(*
SPDX-FileCopyrightText: © 2026 Oleksandr Tiutyk <trofimich@gmail.com>
SPDX-License-Identifier: MIT
License: https://opensource.org/license/mit
*)

(*!
<summary>
Defines a loop composite activity that repeats its body activity while its Condition evaluates to TRUE.
</summary>
*)

INTERFACE IWhileActivity EXTENDS IExclusiveCompositeActivity

(*!
<summary>Returns the body activity executed by this loop, or 0 when no body is configured.</summary>
*)
{attribute 'monitoring' := 'call'}
PROPERTY Body : IActivity
GET
END_GET
END_PROPERTY

(*!
<summary>Returns the loop continuation condition configured for this activity.</summary>
*)
{attribute 'monitoring' := 'call'}
PROPERTY Condition : ICondition
GET
END_GET
END_PROPERTY

(*!
<summary>Configures the required loop condition and optional body activity.</summary>
<description>
Permitted only in PASSIVE_READY. Condition is required; body is optional (when 0, evaluates condition
cyclically without advancing a body activity). Assigns THIS^ as ParentActivity of supplied elements.
</description>
<param name="condition">Condition evaluated before each iteration.</param>
<param name="body">Activity executed repeatedly while condition evaluates to TRUE, or 0.</param>
*)
METHOD Configure
VAR_INPUT
	condition : ICondition;
	body : IActivity;
END_VAR
END_METHOD

END_INTERFACE

(* stored: Version 1.1.0.1
   Itf IWhileActivity: Id {48afd1de-38c9-486e-a527-23b68379f379}
   Property Body: Id {b5e98de3-41de-46f4-b227-f9a8b9545985}
   Get Get: Id {fdec2897-ad2d-4267-821c-cd9a495ee9b5}
   Property Condition: Id {121e9e17-db69-4d58-a344-e6e8a3a42d4b}
   Get Get: Id {9c48afd2-d45d-4366-84e1-f61bd2c6adc9}
   Method Configure: Id {1073bb11-2516-4e4a-b056-d98e3143c9fd} *)
